Fanuc KAREL source: kt00028.KL

-- PROVISIONAL review KL for V770-1; original PC SHA256 0c0f2f1dcc9da9dafe9d40b9aef6e0c047e9fd78ffb24a9b7f12964379949662
-- Incomplete behavior may be omitted. Consult companion uncertainty JSON. Do not deploy.
PROGRAM KT00028
%NOLOCKGROUP
VAR
  R2 : REAL
  OUT : REAL
-- UNRESOLVED_DECL H1 type=002017
BEGIN
  -- UNRESOLVED_PC offsets 5-19; opcodes 2E,22,9D,33,B4
  -- UNRESOLVED_PC offsets 24-35; opcodes 2E,23
  -- UNRESOLVED_PC offsets 40-64; opcodes 22,9D,33,B3,21,29,64,69,23
  -- UNRESOLVED_PC offsets 69-73; opcodes 7F
END KT00028
